// TIA Portal V21 export
// export: Created 2026-10-23T20:44:35.1418135Z, ExportSetting WithDefaults, DisplayName Totally Integrated Automation Portal, DisplayVersion V21 Update 1, DisplayName SINAMICS Startdrive Advanced, DisplayVersion V21 HF2, DisplayName SINAMICS Startdrive G110M, G120, G120C, G120D, G120P, G115D, DisplayVersion V21 HF2, DisplayName SINAMICS Startdrive G130, G150, S120, S150, G200, G220, S200, S210, S220, Innomotics MVD, DisplayVersion V21 HF2, DisplayName STEP 7 Professional, DisplayVersion V21 Update 1, DisplayName STEP 7 Safety, DisplayVersion V21, DisplayName Tech WebApplication, DisplayVersion V21, DisplayName WinCC Basic/Comfort/Advanced, DisplayVersion V21 Update 1, DisplayName WinCC Unified, DisplayVersion V21 Update 1
FUNCTION_BLOCK "FB_Filler"   // FB5, SCL
TITLE = Filler
VERSION : 0.1
// Published filler of the filling unit; uses FC_FillHelper, UDT_FillRecipe and the tags of Tags_Filling
// stored: Access Published, AutoNumber true, IsIECCheckEnabled false, IsRetainMemResEnabled false, MemoryReserve 100, Namespace Filling, SetENOAutomatically false, UDAEnableTagReadback false
   VAR_INPUT
      Start : Bool;   // Start filling
      Stop : Bool;   // Stop filling
   END_VAR
   VAR_OUTPUT
      Filling : Bool;   // Valve is open
      Done : Bool;   // Filling time elapsed or level high
   END_VAR
   VAR_IN_OUT
      Recipe : "Filling.UDT_FillRecipe";   // Active recipe
   END_VAR
   VAR
      FillTimer { S7_SetPoint := 'True'} : TON_TIME;   // Maximum filling time
      Active : Bool;   // Filling is active
   END_VAR
   VAR_TEMP
      Volume : Real;   // Volume from the raw flow
   END_VAR
BEGIN

       REGION Command
           IF #Stop THEN
               #Active := FALSE;
           ELSIF #Start THEN
               #Active := TRUE;
           END_IF;
       END_REGION

       REGION Filling
           #Volume := "Filling.FC_FillHelper"(RawFlow := WORD_TO_INT("FillFlowRaw"), Factor := #Recipe.FlowFactor);
           #FillTimer(IN := #Active, PT := #Recipe.FillTime);
           "FillValveOpen" := #Active AND NOT #FillTimer.Q AND NOT "FillLevelHigh";
       END_REGION

       REGION Outputs
           #Filling := "FillValveOpen";
           #Done := #FillTimer.Q OR "FillLevelHigh";
           #Recipe.LastVolume := #Volume;
       END_REGION
END_FUNCTION_BLOCK
